TYPE Gauge_Type: (
PG722B := 0, //Baraton Gauge
IG903 := 1 , //Cold Cathode
PG907 := 2 , //Pirani Gauge
IG909:= 3 , //Hot Cathode
PG925 := 4 ); //MicroPirani Gauge
(* This enumeration should match up with the EDM MUX button on the vacuum gauge expert controls screen *)
END_TYPE

(* stored: Version 1.1.0.1
   DUT Gauge_Type: Id {c777043f-0b38-4846-b2d2-725c1a5388f6} *)
